Staubli VAL3: sCommentIO.pgx

program sCommentIO()
begin
end
